Staubli VAL3: utEvents.pjx

--- utEvents.pjx ---
Parameters version=s8.8.3Cs9_BS1660 stackSize=5000 millimeterUnit=true
Program file=start.pgx
Program file=stop.pgx
Data file=utEvents.dtx

--- utEvents.dtx ---
public bool bClick
public bool bMouseDown
public bool bMouseUp

--- start.pgx ---
program start()
begin
end

--- stop.pgx ---
program stop()
begin
end
